// TIA Portal project "SnideroEmanuelePLCFineModulo" (V19)

(* hardware
DEVICE "S7-1200 station_1"  S7-1200 Station
   slot 0: "Rack_0"  S7-1200 Rack  Rack  V1.0
   slot 1: "PLC_1"  CPU 1212C DC/DC/Rly  6ES7 212-1HE40-0XB0  V4.6
   slot 2: "DQ 8x24VDC _1"  SM 1222 DQ8 x 24VDC  6ES7 222-1BF32-0XB0  V2.0
DEVICE "HMI_1"  KTP900 Basic PN
   slot 0: "HMI_1"  KTP900 Basic PN  6AV2 123-2JB03-0AX0  17.0.0.0
   slot 1: "HMI_RT_1"  KTP900 Basic PN  6AV2 123-2JB03-0AX0  17.0.0.0
   slot 5: "HMI_1.IE_CP_1"  PROFINET Interface  17.0.0.0
      slot 1: "PROFINET Interface_1"  PROFINET Interface
         slot 1: "Port_1"  Port
*)

// ===== PLC "PLC_1"  CPU 1212C DC/DC/Rly =====

VAR_GLOBAL   // PLC tag table "Default tag table"
   "FotocellulaInserimentoMoneta1Euro" AT %I0.0 : Bool;
   "FotocellulaInserimentoMoneta2Euro" AT %I0.1 : Bool;   // Se un motociclista la inserisce può passare ugualmente, pur senza ricevere resto
   "PlaccaA" AT %I0.2 : Bool;
   "PlaccaB" AT %I0.3 : Bool;
   "PlaccaC" AT %I0.4 : Bool;
   "PlaccaD" AT %I0.5 : Bool;
   "LEDPostiAutoEsauriti" AT %Q0.0 : Bool;
   "LEDPostiMotoEsauriti" AT %Q0.1 : Bool;
   "TeleruttoreS1Su" AT %Q0.2 : Bool;
   "TeleruttoreS1Giù" AT %Q0.3 : Bool;
   "TeleruttoreD1Su" AT %Q0.4 : Bool;
   "TeleruttoreD1Giù" AT %Q0.5 : Bool;
   "TeleruttoreS2Su" AT %Q0.6 : Bool;
   "TeleruttoreS2giù" AT %Q0.7 : Bool;
   "TeleruttoreD2Su" AT %Q1.0 : Bool;
   "TeleruttoreD2Giù" AT %Q1.1 : Bool;
   "AppoggioMoneta1Euro" AT %M0.0 : Bool;
   "AppoggioMoneta2Euro" AT %M0.1 : Bool;
   "AppoggioTeleruttoreS1Su" AT %M0.2 : Bool;
   "AppoggioTeleruttoreD2Su" AT %M0.3 : Bool;
   "AppoggioTeleruttoreD1Su" AT %M0.4 : Bool;
   "Credito" AT %MB10 : SInt;   // Sufficiente credito max 127 euro
   "ResetCreditoManuale" AT %I0.6 : Bool;
   "AppoggioNTeleruttoreS1Su" AT %M0.5 : Bool;
   "AppoggioNQTPS1Sollevata" AT %M0.6 : Bool;
   "AppoggioNTeleruttoreD1Su" AT %M0.7 : Bool;
   "AppoggioNTeleruttoreS2Su" AT %M1.0 : Bool;
   "AppoggioNTeleruttoreD2Su" AT %M1.1 : Bool;
   "AppoggioNQTPD1Sollevata" AT %M1.2 : Bool;
   "AppoggioNQTPS2Sollevata" AT %M1.3 : Bool;
   "AppoggioNQTPD2Sollevata" AT %M1.4 : Bool;
   "AppoggioNQTPS1Discriminazione" AT %M1.5 : Bool;
   "AppoggioNQTPS2Discriminazione" AT %M1.6 : Bool;
   "AppoggioPlaccaA" AT %M1.7 : Bool;
   "AppoggioPlaccaD" AT %M2.0 : Bool;
   "AppoggioTeleruttoreD1SuPostiAuto" AT %M2.1 : Bool;
   "AppoggioTeleruttoreS1SuPostiMoto" AT %M2.2 : Bool;
   "AppoggioTeleruttoreS2Su" AT %Q1.2 : Bool;
   "SelettoreCDAuto" AT %M2.3 : Bool;
   "SelettoreCDMoto" AT %M2.4 : Bool;
   "System_Byte" AT %MB50 : Byte;
   "FirstScan" AT %M50.0 : Bool;
   "DiagStatusUpdate" AT %M50.1 : Bool;
   "AlwaysTRUE" AT %M50.2 : Bool;
   "AlwaysFALSE" AT %M50.3 : Bool;
   "PlaccaAHMI" AT %M2.5 : Bool;
   "PlaccaBHMI" AT %M3.0 : Bool;
   "PlaccaCHMI" AT %M2.7 : Bool;
   "PlaccaDHMI" AT %M2.6 : Bool;
   "FotocellulaInserimentoMoneta1HMI" AT %M3.1 : Bool;
   "FotocellulaInserimentoMoneta2HMI" AT %M3.2 : Bool;
   "ResetCreditoManualeHMI" AT %M3.3 : Bool;
   "AppoggioPlaccaAHMI" AT %M3.4 : Bool;
   "AppoggioPlaccaDHMI" AT %M3.5 : Bool;
   "AppoggioFotocellulaInserimentoMoneta1HMI" AT %M3.6 : Bool;
   "AppoggioFotocellulaInserimentoMoneta2HMI" AT %M3.7 : Bool;
END_VAR

// folder: System blocks/Program resources

DATA_BLOCK "TSalitaS1"   // DB2
{ S7_Optimized_Access := 'TRUE' }
AUTHOR : Simatic
FAMILY : IEC
NAME : IEC_TMR
VERSION : 1.0
// stored: InstanceOfName IEC_TIMER
"IEC_TIMER"
BEGIN
END_DATA_BLOCK

DATA_BLOCK "TDiscesaS1"   // DB3
{ S7_Optimized_Access := 'TRUE' }
AUTHOR : Simatic
FAMILY : IEC
NAME : IEC_TMR
VERSION : 1.0
// stored: InstanceOfName IEC_TIMER
"IEC_TIMER"
BEGIN
END_DATA_BLOCK

DATA_BLOCK "TSalitaD1"   // DB4
{ S7_Optimized_Access := 'TRUE' }
AUTHOR : Simatic
FAMILY : IEC
NAME : IEC_TMR
VERSION : 1.0
// stored: InstanceOfName IEC_TIMER
"IEC_TIMER"
BEGIN
END_DATA_BLOCK

DATA_BLOCK "TDiscesaD1"   // DB5
{ S7_Optimized_Access := 'TRUE' }
AUTHOR : Simatic
FAMILY : IEC
NAME : IEC_TMR
VERSION : 1.0
// stored: InstanceOfName IEC_TIMER
"IEC_TIMER"
BEGIN
END_DATA_BLOCK

DATA_BLOCK "TsalitaS2"   // DB6
{ S7_Optimized_Access := 'TRUE' }
AUTHOR : Simatic
FAMILY : IEC
NAME : IEC_TMR
VERSION : 1.0
// stored: InstanceOfName IEC_TIMER
"IEC_TIMER"
BEGIN
END_DATA_BLOCK

DATA_BLOCK "TDiscesaS2"   // DB7
{ S7_Optimized_Access := 'TRUE' }
AUTHOR : Simatic
FAMILY : IEC
NAME : IEC_TMR
VERSION : 1.0
// stored: InstanceOfName IEC_TIMER
"IEC_TIMER"
BEGIN
END_DATA_BLOCK

DATA_BLOCK "TSalitaD2"   // DB8
{ S7_Optimized_Access := 'TRUE' }
AUTHOR : Simatic
FAMILY : IEC
NAME : IEC_TMR
VERSION : 1.0
// stored: InstanceOfName IEC_TIMER
"IEC_TIMER"
BEGIN
END_DATA_BLOCK

DATA_BLOCK "TDiscesaD2"   // DB9
{ S7_Optimized_Access := 'TRUE' }
AUTHOR : Simatic
FAMILY : IEC
NAME : IEC_TMR
VERSION : 1.0
// stored: InstanceOfName IEC_TIMER
"IEC_TIMER"
BEGIN
END_DATA_BLOCK

DATA_BLOCK "TS1Sollevata"   // DB10
{ S7_Optimized_Access := 'TRUE' }
AUTHOR : Simatic
FAMILY : IEC
NAME : IEC_TMR
VERSION : 1.0
// stored: InstanceOfName IEC_TIMER
"IEC_TIMER"
BEGIN
END_DATA_BLOCK

DATA_BLOCK "TD1Sollevata"   // DB11
{ S7_Optimized_Access := 'TRUE' }
AUTHOR : Simatic
FAMILY : IEC
NAME : IEC_TMR
VERSION : 1.0
// stored: InstanceOfName IEC_TIMER
"IEC_TIMER"
BEGIN
END_DATA_BLOCK

DATA_BLOCK "TS2Sollevata"   // DB12
{ S7_Optimized_Access := 'TRUE' }
AUTHOR : Simatic
FAMILY : IEC
NAME : IEC_TMR
VERSION : 1.0
// stored: InstanceOfName IEC_TIMER
"IEC_TIMER"
BEGIN
END_DATA_BLOCK

DATA_BLOCK "TD2Sollevata"   // DB13
{ S7_Optimized_Access := 'TRUE' }
AUTHOR : Simatic
FAMILY : IEC
NAME : IEC_TMR
VERSION : 1.0
// stored: InstanceOfName IEC_TIMER
"IEC_TIMER"
BEGIN
END_DATA_BLOCK

DATA_BLOCK "CTUDAuto"   // DB14
{ S7_Optimized_Access := 'TRUE' }
AUTHOR : Simatic
FAMILY : IEC
NAME : CNTR
VERSION : 1.0
// stored: InstanceOfName IEC_COUNTER
"IEC_COUNTER"
BEGIN
END_DATA_BLOCK

DATA_BLOCK "CTUDMoto"   // DB15
{ S7_Optimized_Access := 'TRUE' }
AUTHOR : Simatic
FAMILY : IEC
NAME : CNTR
VERSION : 1.0
// stored: InstanceOfName IEC_COUNTER
"IEC_COUNTER"
BEGIN
END_DATA_BLOCK

DATA_BLOCK "TPS1DiscriminazioneMezzo"   // DB17
{ S7_Optimized_Access := 'TRUE' }
AUTHOR : Simatic
FAMILY : IEC
NAME : IEC_TMR
VERSION : 1.0
// stored: InstanceOfName IEC_TIMER
"IEC_TIMER"
BEGIN
END_DATA_BLOCK

DATA_BLOCK "TPS2DiscriminazioneMezzo"   // DB18
{ S7_Optimized_Access := 'TRUE' }
AUTHOR : Simatic
FAMILY : IEC
NAME : IEC_TMR
VERSION : 1.0
// stored: InstanceOfName IEC_TIMER
"IEC_TIMER"
BEGIN
END_DATA_BLOCK

// folder: (top level)

ORGANIZATION_BLOCK "Main"   // OB1, LAD, ProgramCycle
TITLE = "Main Program Sweep (Cycle)"
{ S7_Optimized_Access := 'TRUE' }
VERSION : 0.1
   VAR_INPUT
      Initial_Call : Bool;   // Initial call of this OB
      Remanence : Bool;   // =True, if remanent data are available
   END_VAR
   VAR_TEMP   // added for the SCL form of the ladder/FBD networks
      _w1 : Bool;
      _w2 : Bool;
      _w3 : Bool;
      _w4 : Bool;
      _w5 : Bool;
      _w6 : Bool;
   END_VAR
BEGIN

REGION Network 1
   // Conteggio monete
   // Le due gettoniere hanno serbatoio in comune.
   // Il conteggio tiene conto del credito (NON MONETE, dunque) totale disponibile
   // 
   // Siccome è possibile inserire monete anche quando nessun mezzo è posizionato sulle placche, il serbatoio delle gettoniere non ha limiti (max 127, comunque. Poi toccherebbe a un operatore svuotare il serbatoio e azzerare il credito manualmente...).
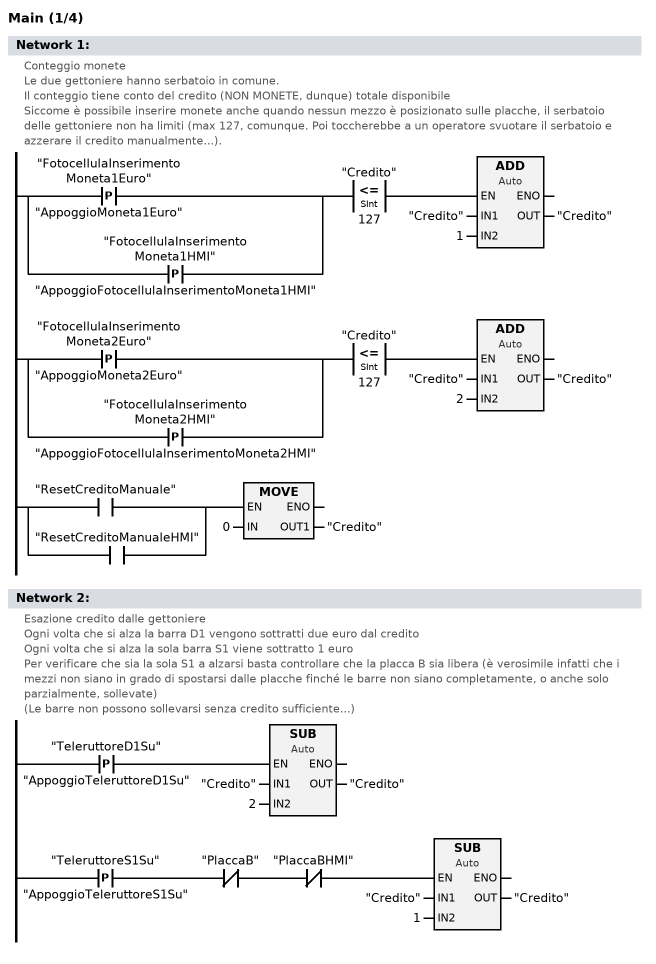
   RUNG wire#powerrail
      P_Contact(operand := "FotocellulaInserimentoMoneta1Euro", bit := "AppoggioMoneta1Euro")
      wire#w1
      { S7_Templates := "SrcType := SInt" } LE_Contact(in1 := "Credito", in2 := 127)
      Add(in1 := "Credito", in2 := 1, out => "Credito")
   END_RUNG
   RUNG wire#powerrail
      P_Contact(operand := "FotocellulaInserimentoMoneta1HMI", bit := "AppoggioFotocellulaInserimentoMoneta1HMI")
   END_RUNG wire#w1
   RUNG wire#powerrail
      P_Contact(operand := "FotocellulaInserimentoMoneta2Euro", bit := "AppoggioMoneta2Euro")
      wire#w2
      { S7_Templates := "SrcType := SInt" } LE_Contact(in1 := "Credito", in2 := 127)
      Add(in1 := "Credito", in2 := 2, out => "Credito")
   END_RUNG
   RUNG wire#powerrail
      P_Contact(operand := "FotocellulaInserimentoMoneta2HMI", bit := "AppoggioFotocellulaInserimentoMoneta2HMI")
   END_RUNG wire#w2
   RUNG wire#powerrail
      Contact( "ResetCreditoManuale" )
      wire#w3
      Move(in := 0, out1 => "Credito")
   END_RUNG
   RUNG wire#powerrail
      Contact( "ResetCreditoManualeHMI" )
   END_RUNG wire#w3
   // the same network as SCL:
   #_w1 := "FotocellulaInserimentoMoneta1Euro" AND NOT "AppoggioMoneta1Euro";   // rising edge of "FotocellulaInserimentoMoneta1Euro"
   "AppoggioMoneta1Euro" := "FotocellulaInserimentoMoneta1Euro";
   #_w2 := "FotocellulaInserimentoMoneta1HMI" AND NOT "AppoggioFotocellulaInserimentoMoneta1HMI";   // rising edge of "FotocellulaInserimentoMoneta1HMI"
   "AppoggioFotocellulaInserimentoMoneta1HMI" := "FotocellulaInserimentoMoneta1HMI";
   IF (#_w1 OR #_w2) AND ("Credito" <= 127) THEN "Credito" := "Credito" + 1; END_IF;
   #_w3 := "FotocellulaInserimentoMoneta2Euro" AND NOT "AppoggioMoneta2Euro";   // rising edge of "FotocellulaInserimentoMoneta2Euro"
   "AppoggioMoneta2Euro" := "FotocellulaInserimentoMoneta2Euro";
   #_w4 := "FotocellulaInserimentoMoneta2HMI" AND NOT "AppoggioFotocellulaInserimentoMoneta2HMI";   // rising edge of "FotocellulaInserimentoMoneta2HMI"
   "AppoggioFotocellulaInserimentoMoneta2HMI" := "FotocellulaInserimentoMoneta2HMI";
   IF (#_w3 OR #_w4) AND ("Credito" <= 127) THEN "Credito" := "Credito" + 2; END_IF;
   IF "ResetCreditoManuale" OR "ResetCreditoManualeHMI" THEN "Credito" := 0; END_IF;
END_REGION

REGION Network 2
   // Esazione credito dalle gettoniere
   // 
   // Ogni volta che si alza la barra D1 vengono sottratti due euro dal credito
   // 
   // Ogni volta che si alza la sola barra S1 viene sottratto 1 euro
   // Per verificare che sia la sola S1 a alzarsi basta controllare che la placca B sia libera (è verosimile infatti che i mezzi non siano in grado di spostarsi dalle placche finché le barre non siano completamente, o anche solo parzialmente, sollevate)
   // 
   // (Le barre non possono sollevarsi senza credito sufficiente...)
   RUNG wire#powerrail
      P_Contact(operand := "TeleruttoreD1Su", bit := "AppoggioTeleruttoreD1Su")
      Sub(in1 := "Credito", in2 := 2, out => "Credito")
   END_RUNG
   RUNG wire#powerrail
      P_Contact(operand := "TeleruttoreS1Su", bit := "AppoggioTeleruttoreS1Su")
      I_Contact( "PlaccaB" )
      I_Contact( "PlaccaBHMI" )
      Sub(in1 := "Credito", in2 := 1, out => "Credito")
   END_RUNG
   // the same network as SCL:
   #_w1 := "TeleruttoreD1Su" AND NOT "AppoggioTeleruttoreD1Su";   // rising edge of "TeleruttoreD1Su"
   "AppoggioTeleruttoreD1Su" := "TeleruttoreD1Su";
   IF #_w1 THEN "Credito" := "Credito" - 2; END_IF;
   #_w2 := "TeleruttoreS1Su" AND NOT "AppoggioTeleruttoreS1Su";   // rising edge of "TeleruttoreS1Su"
   "AppoggioTeleruttoreS1Su" := "TeleruttoreS1Su";
   IF #_w2 AND NOT "PlaccaB" AND NOT "PlaccaBHMI" THEN "Credito" := "Credito" - 1; END_IF;
END_REGION

REGION Network 3
   // Barra S1
   // 
   // Non può alzarsi se 
   // - i posti moto occupati sono già 8 (e la sola placca A è attiva) o non vi è credito disponibile maggiore o uguale a 1
   // - i posti auto occupati sono già 8 (e entrambe le placche sono attive) o non vi è credito disponibile maggiore o uguale a 2
   // - è ancora in stato di sosta in alto o di discesa
   // 
   // Se entro 2 secondi dall'attivazione della placca A non si attiva anche la B il veicolo viene considerato una moto.
   // 
   // La durata della sosta alzata viene aggiornata quando la barra si è completamente alzata, sulla base delle placche attive in quel momento (si considera che i mezzi non possano spostarsi da esse finché le barre non sono completamente alzate)
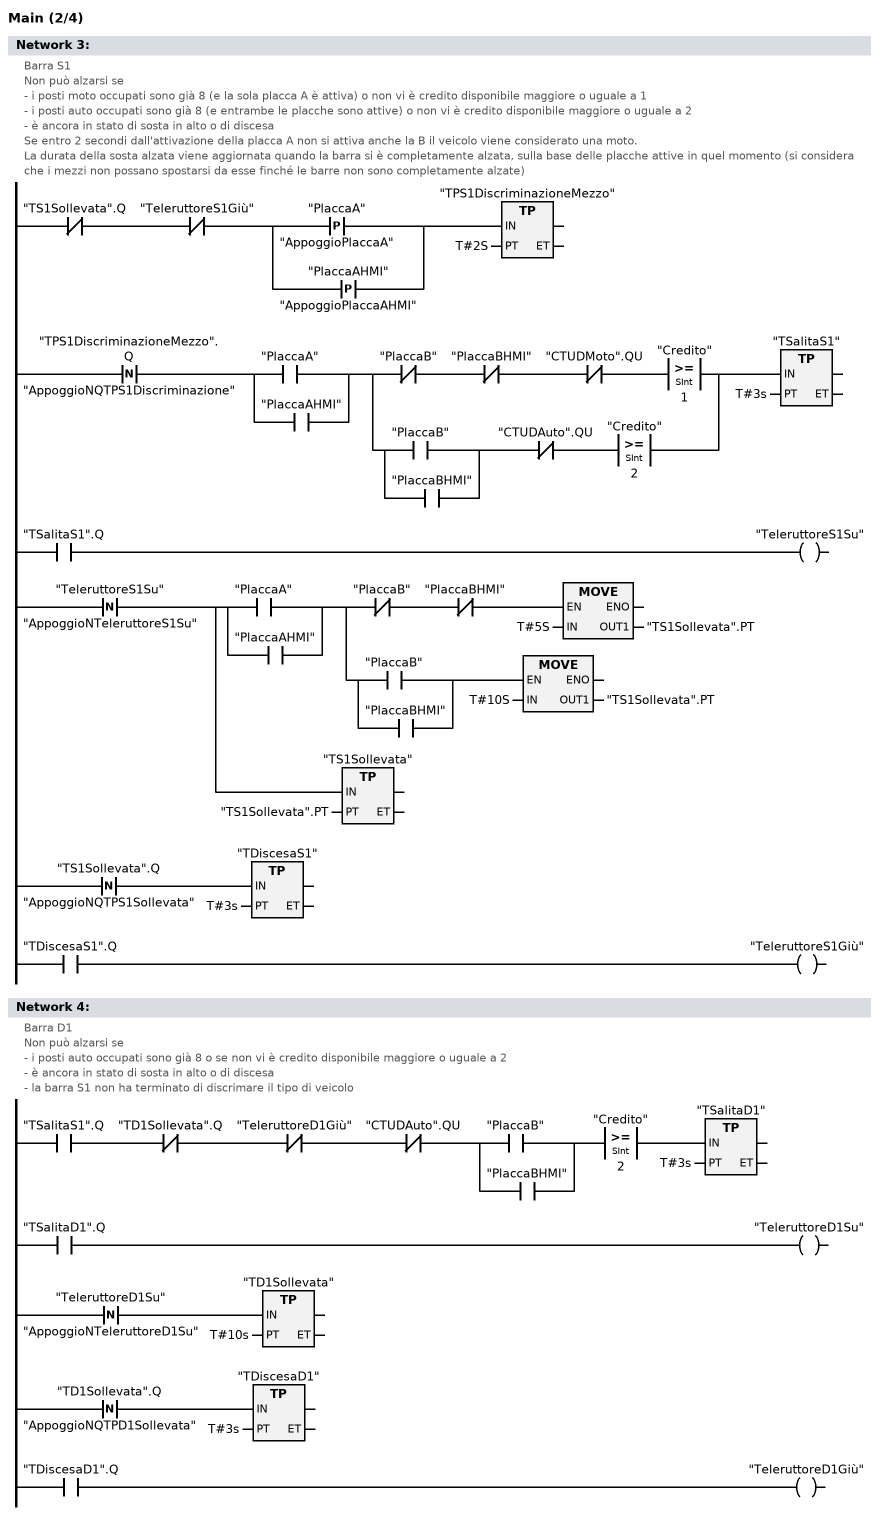
   #_w1 := NOT "TS1Sollevata".Q AND NOT "TeleruttoreS1Giù" AND "PlaccaA" AND NOT "AppoggioPlaccaA";   // rising edge of "PlaccaA"
   "AppoggioPlaccaA" := "PlaccaA";
   #_w2 := NOT "TS1Sollevata".Q AND NOT "TeleruttoreS1Giù" AND "PlaccaAHMI" AND NOT "AppoggioPlaccaAHMI";   // rising edge of "PlaccaAHMI"
   "AppoggioPlaccaAHMI" := "PlaccaAHMI";
   "TPS1DiscriminazioneMezzo".TP(IN := #_w1 OR #_w2, PT := T#2S);
   #_w3 := NOT "TPS1DiscriminazioneMezzo".Q AND "AppoggioNQTPS1Discriminazione";   // falling edge of "TPS1DiscriminazioneMezzo".Q
   "AppoggioNQTPS1Discriminazione" := "TPS1DiscriminazioneMezzo".Q;
   "TSalitaS1".TP(IN := #_w3 AND ("PlaccaA" OR "PlaccaAHMI") AND ((NOT "PlaccaB" AND NOT "PlaccaBHMI" AND NOT "CTUDMoto".QU AND ("Credito" >= 1)) OR (("PlaccaB" OR "PlaccaBHMI") AND NOT "CTUDAuto".QU AND ("Credito" >= 2))),
                  PT := T#3s);
   "TeleruttoreS1Su" := "TSalitaS1".Q;
   #_w4 := NOT "TeleruttoreS1Su" AND "AppoggioNTeleruttoreS1Su";   // falling edge of "TeleruttoreS1Su"
   "AppoggioNTeleruttoreS1Su" := "TeleruttoreS1Su";
   #_w5 := #_w4 AND ("PlaccaA" OR "PlaccaAHMI");
   IF #_w5 AND NOT "PlaccaB" AND NOT "PlaccaBHMI" THEN "TS1Sollevata".PT := T#5S; END_IF;
   IF #_w5 AND ("PlaccaB" OR "PlaccaBHMI") THEN "TS1Sollevata".PT := T#10S; END_IF;
   "TS1Sollevata".TP(IN := #_w4, PT := "TS1Sollevata".PT);
   #_w6 := NOT "TS1Sollevata".Q AND "AppoggioNQTPS1Sollevata";   // falling edge of "TS1Sollevata".Q
   "AppoggioNQTPS1Sollevata" := "TS1Sollevata".Q;
   "TDiscesaS1".TP(IN := #_w6, PT := T#3s);
   "TeleruttoreS1Giù" := "TDiscesaS1".Q;
END_REGION

REGION Network 4
   // Barra D1
   // 
   // Non può alzarsi se
   // - i posti auto occupati sono già 8 o se non vi è credito disponibile maggiore o uguale a 2
   // - è ancora in stato di sosta in alto o di discesa
   // - la barra S1 non ha terminato di discrimare il tipo di veicolo
   "TSalitaD1".TP(IN := "TSalitaS1".Q AND NOT "TD1Sollevata".Q AND NOT "TeleruttoreD1Giù" AND NOT "CTUDAuto".QU AND ("PlaccaB" OR "PlaccaBHMI") AND ("Credito" >= 2),
                  PT := T#3s);
   "TeleruttoreD1Su" := "TSalitaD1".Q;
   #_w1 := NOT "TeleruttoreD1Su" AND "AppoggioNTeleruttoreD1Su";   // falling edge of "TeleruttoreD1Su"
   "AppoggioNTeleruttoreD1Su" := "TeleruttoreD1Su";
   "TD1Sollevata".TP(IN := #_w1, PT := T#10s);
   #_w2 := NOT "TD1Sollevata".Q AND "AppoggioNQTPD1Sollevata";   // falling edge of "TD1Sollevata".Q
   "AppoggioNQTPD1Sollevata" := "TD1Sollevata".Q;
   "TDiscesaD1".TP(IN := #_w2, PT := T#3s);
   "TeleruttoreD1Giù" := "TDiscesaD1".Q;
END_REGION

REGION Network 5
   // Barra S2
   // 
   // Sufficiente sia attiva la placca D perchè si alzi.
   // 
   // Per permettere all'eventuale auto di piazzarsi anche sulla C vengono concessi 2 secondi
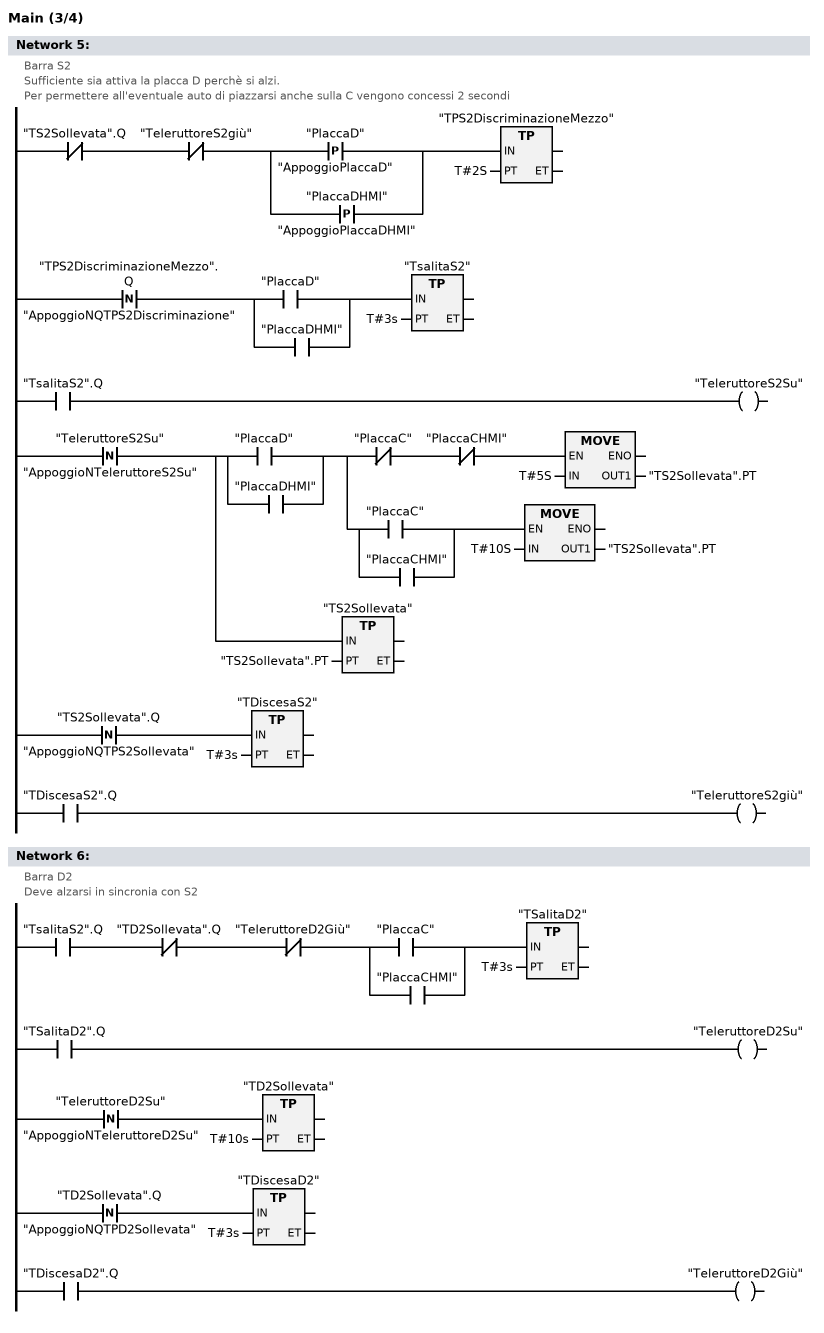
   #_w1 := NOT "TS2Sollevata".Q AND NOT "TeleruttoreS2giù" AND "PlaccaD" AND NOT "AppoggioPlaccaD";   // rising edge of "PlaccaD"
   "AppoggioPlaccaD" := "PlaccaD";
   #_w2 := NOT "TS2Sollevata".Q AND NOT "TeleruttoreS2giù" AND "PlaccaDHMI" AND NOT "AppoggioPlaccaDHMI";   // rising edge of "PlaccaDHMI"
   "AppoggioPlaccaDHMI" := "PlaccaDHMI";
   "TPS2DiscriminazioneMezzo".TP(IN := #_w1 OR #_w2, PT := T#2S);
   #_w3 := NOT "TPS2DiscriminazioneMezzo".Q AND "AppoggioNQTPS2Discriminazione";   // falling edge of "TPS2DiscriminazioneMezzo".Q
   "AppoggioNQTPS2Discriminazione" := "TPS2DiscriminazioneMezzo".Q;
   "TsalitaS2".TP(IN := #_w3 AND ("PlaccaD" OR "PlaccaDHMI"), PT := T#3s);
   "TeleruttoreS2Su" := "TsalitaS2".Q;
   #_w4 := NOT "TeleruttoreS2Su" AND "AppoggioNTeleruttoreS2Su";   // falling edge of "TeleruttoreS2Su"
   "AppoggioNTeleruttoreS2Su" := "TeleruttoreS2Su";
   #_w5 := #_w4 AND ("PlaccaD" OR "PlaccaDHMI");
   IF #_w5 AND NOT "PlaccaC" AND NOT "PlaccaCHMI" THEN "TS2Sollevata".PT := T#5S; END_IF;
   IF #_w5 AND ("PlaccaC" OR "PlaccaCHMI") THEN "TS2Sollevata".PT := T#10S; END_IF;
   "TS2Sollevata".TP(IN := #_w4, PT := "TS2Sollevata".PT);
   #_w6 := NOT "TS2Sollevata".Q AND "AppoggioNQTPS2Sollevata";   // falling edge of "TS2Sollevata".Q
   "AppoggioNQTPS2Sollevata" := "TS2Sollevata".Q;
   "TDiscesaS2".TP(IN := #_w6, PT := T#3s);
   "TeleruttoreS2giù" := "TDiscesaS2".Q;
END_REGION

REGION Network 6
   // Barra D2
   // 
   // Deve alzarsi in sincronia con S2
   "TSalitaD2".TP(IN := "TsalitaS2".Q AND NOT "TD2Sollevata".Q AND NOT "TeleruttoreD2Giù" AND ("PlaccaC" OR "PlaccaCHMI"),
                  PT := T#3s);
   "TeleruttoreD2Su" := "TSalitaD2".Q;
   #_w1 := NOT "TeleruttoreD2Su" AND "AppoggioNTeleruttoreD2Su";   // falling edge of "TeleruttoreD2Su"
   "AppoggioNTeleruttoreD2Su" := "TeleruttoreD2Su";
   "TD2Sollevata".TP(IN := #_w1, PT := T#10s);
   #_w2 := NOT "TD2Sollevata".Q AND "AppoggioNQTPD2Sollevata";   // falling edge of "TD2Sollevata".Q
   "AppoggioNQTPD2Sollevata" := "TD2Sollevata".Q;
   "TDiscesaD2".TP(IN := #_w2, PT := T#3s);
   "TeleruttoreD2Giù" := "TDiscesaD2".Q;
END_REGION

REGION Network 7
   // Ogni volta che si alza la barra D1 (non può alzarsi quando 8 posti sono già occupati) il conteggio incrementa
   // Quando si alza la D2 decrementa
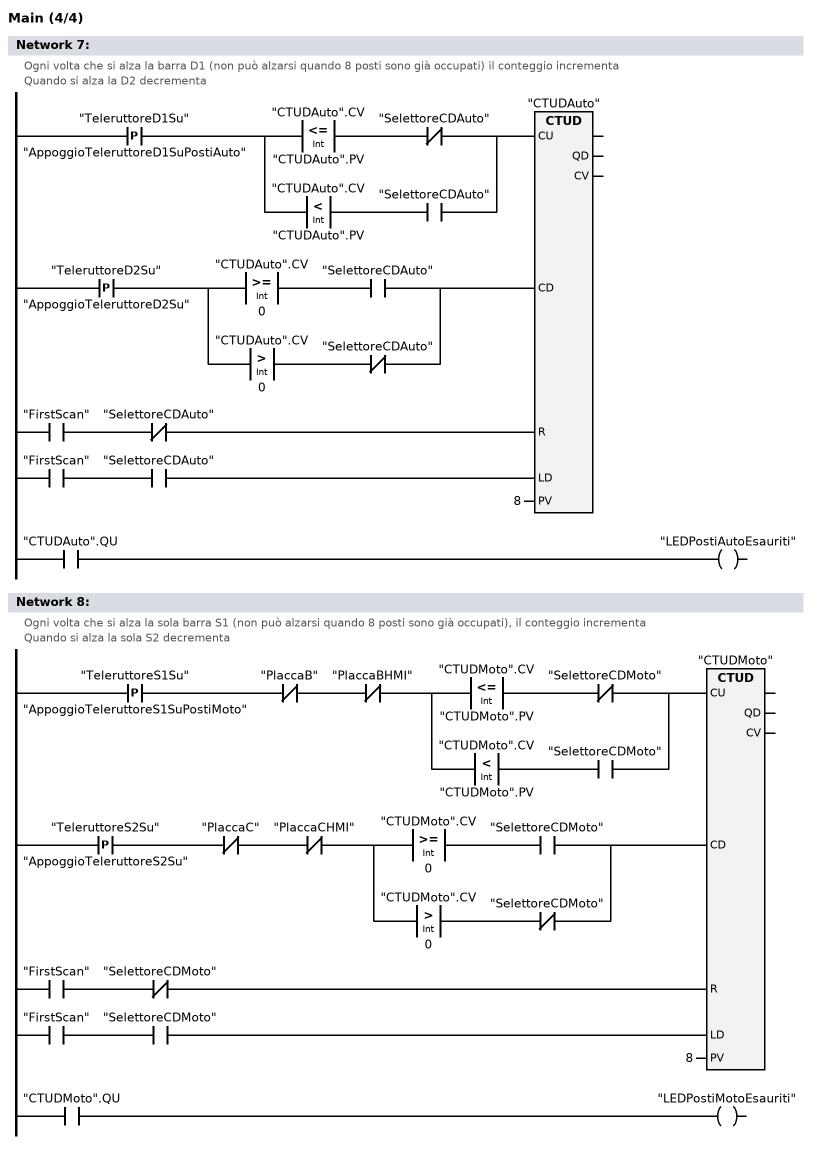
   #_w1 := "TeleruttoreD1Su" AND NOT "AppoggioTeleruttoreD1SuPostiAuto";   // rising edge of "TeleruttoreD1Su"
   "AppoggioTeleruttoreD1SuPostiAuto" := "TeleruttoreD1Su";
   #_w2 := "TeleruttoreD2Su" AND NOT "AppoggioTeleruttoreD2Su";   // rising edge of "TeleruttoreD2Su"
   "AppoggioTeleruttoreD2Su" := "TeleruttoreD2Su";
   "CTUDAuto".CTUD(CU := #_w1 AND ((("CTUDAuto".CV <= "CTUDAuto".PV) AND NOT "SelettoreCDAuto") OR (("CTUDAuto".CV < "CTUDAuto".PV) AND "SelettoreCDAuto")),
                   CD := #_w2 AND ((("CTUDAuto".CV >= 0) AND "SelettoreCDAuto") OR (("CTUDAuto".CV > 0) AND NOT "SelettoreCDAuto")),
                   R := "FirstScan" AND NOT "SelettoreCDAuto",
                   LD := "FirstScan" AND "SelettoreCDAuto",
                   PV := 8);
   "LEDPostiAutoEsauriti" := "CTUDAuto".QU;
END_REGION

REGION Network 8
   // Ogni volta che si alza la sola barra S1 (non può alzarsi quando 8 posti sono già occupati), il conteggio incrementa
   // Quando si alza la sola S2 decrementa
   #_w1 := "TeleruttoreS1Su" AND NOT "AppoggioTeleruttoreS1SuPostiMoto";   // rising edge of "TeleruttoreS1Su"
   "AppoggioTeleruttoreS1SuPostiMoto" := "TeleruttoreS1Su";
   #_w2 := "TeleruttoreS2Su" AND NOT "AppoggioTeleruttoreS2Su";   // rising edge of "TeleruttoreS2Su"
   "AppoggioTeleruttoreS2Su" := "TeleruttoreS2Su";
   "CTUDMoto".CTUD(CU := #_w1 AND NOT "PlaccaB" AND NOT "PlaccaBHMI" AND ((("CTUDMoto".CV <= "CTUDMoto".PV) AND NOT "SelettoreCDMoto") OR (("CTUDMoto".CV < "CTUDMoto".PV) AND "SelettoreCDMoto")),
                   CD := #_w2 AND NOT "PlaccaC" AND NOT "PlaccaCHMI" AND ((("CTUDMoto".CV >= 0) AND "SelettoreCDMoto") OR (("CTUDMoto".CV > 0) AND NOT "SelettoreCDMoto")),
                   R := "FirstScan" AND NOT "SelettoreCDMoto",
                   LD := "FirstScan" AND "SelettoreCDMoto",
                   PV := 8);
   "LEDPostiMotoEsauriti" := "CTUDMoto".QU;
END_REGION
END_ORGANIZATION_BLOCK

(* ===== HMI "HMI_RT_1" =====
system functions are stored by id; their names below are inferred from use
connection "HMI_Connection_1": ETHERNET, SMART_S7_1200_OMS

HMI tags "Default tag table"
   "Tag_ScreenNumber" : UInt, internal
   "PlaccaAHMI" : Bool = PLC PlaccaAHMI AT %M2.5, 100 ms
   "PlaccaBHMI" : Bool = PLC PlaccaBHMI AT %M3.0, 100 ms
   "PlaccaCHMI" : Bool = PLC PlaccaCHMI AT %M2.7, 100 ms
   "PlaccaDHMI" : Bool = PLC PlaccaDHMI AT %M2.6, 100 ms
   "ResetCreditoManualeHMI" : Bool = PLC ResetCreditoManualeHMI AT %M3.3, 100 ms
   "CTUDMoto_CV" : Int = PLC CTUDMoto.CV, 100 ms
   "CTUDAuto_CV" : Int = PLC CTUDAuto.CV, 100 ms
   "FotocellulaInserimentoMoneta1HMI" : Bool = PLC FotocellulaInserimentoMoneta1HMI AT %M3.1, 100 ms
   "FotocellulaInserimentoMoneta2HMI" : Bool = PLC FotocellulaInserimentoMoneta2HMI AT %M3.2, 100 ms
   "LEDPostiMotoEsauriti" : Bool = PLC LEDPostiMotoEsauriti AT %Q0.1, 100 ms
   "LEDPostiAutoEsauriti" : Bool = PLC LEDPostiAutoEsauriti AT %Q0.0, 100 ms
   "Credito" : SInt = PLC Credito AT %MB10, 100 ms
   "TD1Sollevata_Q" : Bool = PLC TD1Sollevata.Q, 1 s
   "TS1Sollevata_Q" : Bool = PLC TS1Sollevata.Q, 1 s
   "TD2Sollevata_Q" : Bool = PLC TD2Sollevata.Q, 1 s
   "TS2Sollevata_Q" : Bool = PLC TS2Sollevata.Q, 1 s
   "TeleruttoreS1Su" : Bool = PLC TeleruttoreS1Su AT %Q0.2, 1 s

Template "Template_1" 800x480
   Button "Exit" at 722,440 size 55x39; TextOff 'Exit'; PictureOff "ExitRuntime_KTP900_Basic_PN_TR"; PictureOn "ExitRuntime_KTP900_Basic_PN_TR"
      on Release: StopRuntime(0)
   Button "Template_Button" at 622,440 size 55x39; TextOff 'Text'
   Button "Template_Button_1" at 522,440 size 55x39; TextOff 'Text'
   Button "Template_Button_2" at 422,440 size 55x39; TextOff 'Text'
   Button "Template_Button_3" at 322,440 size 55x39; TextOff 'Text'
   Button "Template_Button_4" at 222,440 size 55x39; TextOff 'Text'
   Button "Alarms" at 122,440 size 55x39; TextOff 'Alarms'; PictureOff "AlarmDisplay_KTP900_Basic_PN_TR"; PictureOn "AlarmDisplay_KTP900_Basic_PN_TR"
      on Release: function_ef3f5d25("Alarm window_Unacknowledged", -1)
   Button "Start screen" at 22,440 size 55x39; TextOff 'Start screen'; PictureOff "NavigateHome_KTP900_Basic_PN_TR"; PictureOn "NavigateHome_KTP900_Basic_PN_TR"
      on Release: ActivateScreen("Root screen", 0)
   SymbolicIOField "Symbolic_IO_Field_Screen" at 73,7 size 620x26; TextOff '0'; TextOn '1'; TextList "TextList_ScreenNames"
      ProcessValue <- "Tag_ScreenNumber"
      on Change: ActivateScreenByNumber("Tag_ScreenNumber", 0)
   DateTimeField "HmiScreenItemData" at 695,20 size 105x20
   DateTimeField "HmiScreenItemData_1" at 695,0 size 105x20
   GraphicView "Logo" at 0,0 size 71x40; Picture "Logo of HMI_1"

screen "Root screen" 800x480, template "Template_1"
   on GenerateScreen: SetTag("Tag_ScreenNumber", 1)
   GraphicView "Graphic view_10" at 644,389 size 96x48; Picture "BarraSollevataVert"
      Visibility <- "TS2Sollevata_Q"
   GraphicView "Graphic view_9" at 539,389 size 96x48; Picture "BarraSollevataVertOriz"
      Visibility <- "TD2Sollevata_Q"
   GraphicView "Graphic view_8" at 344,215 size 96x48; Picture "BarraSollevata"
      Visibility <- "TD1Sollevata_Q"
   GraphicView "Graphic view_7" at 238,215 size 96x48; Picture "BarraSollevataOriz"
      Visibility <- "TS1Sollevata_Q"
   GraphicView "Graphic view_6" at 643,385 size 96x48; Picture "BarraVert"
      Visibility <- "TS2Sollevata_Q"
   GraphicView "Graphic view_5" at 542,385 size 96x48; Picture "BarraVertOriz"
      Visibility <- "TD2Sollevata_Q"
   GraphicView "Graphic view_4" at 341,219 size 96x48; Picture "Barra"
      Visibility <- "TD1Sollevata_Q"
   GraphicView "Graphic view_3" at 242,219 size 96x48; Picture "BarraCapovolta"
      Visibility <- "TS1Sollevata_Q"
   TextField "HmiScreenItemData" at 243,114 size 195x28; Text 'PARCHEGGIO'
   GraphicView "Graphic view_1" at 291,238 size 96x198; Picture "Carreggiata"
   GraphicView "Graphic view_2" at 592,219 size 96x196; Picture "Carreggiata"
   Button "FB_ArrowUp_Round" at 343,339 size 43x44; TextOff 'Text'; PictureOff "FB_ArrowUp_Round_Released_256c"; PictureOn "FB_ArrowUp_Round_Pressed_256c"
      on Press: SetBit("PlaccaBHMI")
      on Release: ResetBit("PlaccaBHMI")
   Button "FB_ArrowUp_Round_1" at 291,339 size 43x44; TextOff 'Text'; PictureOff "FB_ArrowUp_Round_Released_256c"; PictureOn "FB_ArrowUp_Round_Pressed_256c"
      on Press: SetBit("PlaccaAHMI")
      on Release: ResetBit("PlaccaAHMI")
   Button "FB_ArrowDown_Round" at 594,256 size 44x46; TextOff 'Text'; PictureOff "FB_ArrowDown_Round_Released_256c"; PictureOn "FB_ArrowDown_Round_Pressed_256c"
      on Press: SetBit("PlaccaCHMI")
      on Release: ResetBit("PlaccaCHMI")
   Button "FB_ArrowDown_Round_1" at 644,256 size 44x46; TextOff 'Text'; PictureOff "FB_ArrowDown_Round_Released_256c"; PictureOn "FB_ArrowDown_Round_Pressed_256c"
      on Press: SetBit("PlaccaDHMI")
      on Release: ResetBit("PlaccaDHMI")
   TextField "Text field_1" at 300,385 size 26x26; Text 'A'
   TextField "Text field_2" at 352,385 size 24x26; Text 'B'
   TextField "Text field_3" at 604,226 size 24x26; Text 'C'
   TextField "Text field_4" at 653,226 size 25x26; Text 'D'
   Button "FB_Attention_Round" at 141,298 size 50x50; TextOff 'Text'; PictureOff "FB_Attention_Round_Released_256c"; PictureOn "FB_Attention_Round_Pressed_256c"
      on Press: SetBit("ResetCreditoManualeHMI")
      on Release: ResetBit("ResetCreditoManualeHMI")
   TextField "Text field_5" at 121,272 size 94x20; Text 'Reset Credito'
   IOField "I/O field_1" at 394,174 size 96x32; FormatPattern 99999
      ProcessValue <- "CTUDAuto_CV"
   IOField "I/O field_2" at 190,174 size 96x32; FormatPattern 99999
      ProcessValue <- "CTUDMoto_CV"
   TextField "HmiScreenItemData_1" at 190,152 size 90x22; Text 'Moto'
   TextField "HmiScreenItemData_2" at 392,151 size 98x22; Text 'Auto'
   TextField "Text field_6" at 17,228 size 82x20; Text 'GETTONIERA'
   TextField "Text field_7" at 58,309 size 21x20; Text '1€'
   TextField "Text field_8" at 58,350 size 21x20; Text '2€'
   Button "FB_ArrowLeft_Round" at 86,308 size 41x37; TextOff 'Text'; PictureOff "FB_ArrowLeft_Round_Released_256c"; PictureOn "FB_ArrowLeft_Round_Pressed_256c"
      on Press: SetBit("FotocellulaInserimentoMoneta1HMI")
      on Release: ResetBit("FotocellulaInserimentoMoneta1HMI")
   Button "FB_ArrowLeft_Round_1" at 86,349 size 40x38; TextOff 'Text'; PictureOff "FB_ArrowLeft_Round_Released_256c"; PictureOn "FB_ArrowLeft_Round_Pressed_256c"
      on Release: ResetBit("FotocellulaInserimentoMoneta2HMI")
      on Press: SetBit("FotocellulaInserimentoMoneta2HMI")
   Circle "Circle_1" at 134,159 size 48x48
      Appearance <- "LEDPostiMotoEsauriti"
   Circle "Circle_2" at 505,159 size 48x48
      Appearance <- "LEDPostiAutoEsauriti"
   IOField "I/O field_3" at 18,267 size 82x32; FormatPattern 999
      ProcessValue <- "Credito"
   TextField "Text field_9" at 35,247 size 52x20; Text 'Credito'
   Button "FB_ArrowUp_Round_2" at 298,245 size 83x50; TextOff 'Text'; PictureOff "FB_ArrowUp_Round_Released_256c"; PictureOn "FB_ArrowUp_Round_Pressed_256c"
      on Press: SetBit("PlaccaAHMI"); SetBit("PlaccaBHMI")
      on Release: ResetBit("PlaccaAHMI"); ResetBit("PlaccaBHMI")
   TextField "Text field_10" at 312,297 size 53x26; Text 'A + B'
   Button "FB_ArrowDown_Round_2" at 600,350 size 80x50; TextOff 'Text'; PictureOff "FB_ArrowDown_Round_Released_256c"; PictureOn "FB_ArrowDown_Round_Pressed_256c"
      on Press: SetBit("PlaccaCHMI"); SetBit("PlaccaDHMI")
      on Release: ResetBit("PlaccaCHMI"); ResetBit("PlaccaDHMI")
   TextField "Text field_11" at 614,321 size 52x26; Text 'C + D'
*)